Fanuc KAREL source: kb00007.KL

-- PROVISIONAL review KL for V770-1; original PC SHA256 1d6e598083e759088f5d322977d0e5cd6439afba7fd8de1f5ad3be010b2e91ea
-- Incomplete behavior may be omitted. Consult companion uncertainty JSON. Do not deploy.
PROGRAM KB00007
%NOLOCKGROUP
BEGIN
  -- UNRESOLVED_PC offsets 5-28; opcodes 27,22,1C,31,4A
  -- UNRESOLVED_PC offsets 33-37; opcodes 7F
END KB00007
